{attribute 'linkalways'} 
{attribute 'no_explicit_call' := 'This FB is a CLASS and must be accessed using methods or properties'}
{attribute 'enable_dynamic_creation'}
FUNCTION_BLOCK  PUBLIC Ax5000 IMPLEMENTS Drive
VAR
END_VAR

END_FUNCTION_BLOCK

(* stored: Version 1.1.0.1
   POU Ax5000: Id {775e59cb-0ef8-4f4c-89b5-46e996c161b8}, SpecialFunc None *)
